FUNCTION_BLOCK FB_AxesEnable
VAR_INPUT
	bEnableAxes: 		BOOL := TRUE;
	bEnableXY:			BOOL;
	bEnableZp:			BOOL;
	bEnableZn:			BOOL;
	bReset:				BOOL;
	fOverride:			LREAL := 10;
END_VAR             	
VAR_OUTPUT          	
	bAllAxesReady:		BOOL := FALSE;
	fbError:			FB_Error;
END_VAR             	
VAR_IN_OUT          	
	stX:				AXIS_REF;
	stY:				AXIS_REF;
	stZ:				AXIS_REF;
END_VAR
VAR	
//Freigaben
	fbPowerX:			MC_Power;
	fbPowerY:			MC_Power;
	fbPowerZ:			MC_Power;
END_VAR


IF NOT (__ISVALIDREF(stX) AND __ISVALIDREF(stY) AND __ISVALIDREF(stZ)) THEN
	fbError.M_Set(1798, 'Üngültige Referenz der Achsen', 0, eID := E_ErrorIDs.eInvalidReference, eSrc := E_ErrorSrcs.ePlc);
	RETURN;
END_IF

IF bReset THEN
	fbError.M_Reset();
	bReset := FALSE;
END_IF

stX.ReadStatus();
stY.ReadStatus();
stZ.ReadStatus();

fbPowerX(
	Enable:=bEnableAxes AND bEnableXY, 
	Enable_Positive:=bEnableAxes AND bEnableXY, 
	Enable_Negative:=bEnableAxes AND bEnableXY, 
	Override:=fOverride, 
	BufferMode:= , 
	Axis:=stX, 
	Status=> , 
	Busy=> , 
	Active=> , 
	Error=> , 
	ErrorID=> );
	
fbPowerY(
	Enable:=bEnableAxes AND bEnableXY, 
	Enable_Positive:=bEnableAxes AND bEnableXY, 
	Enable_Negative:=bEnableAxes AND bEnableXY, 
	Override:=fOverride, 
	BufferMode:= , 
	Axis:=stY, 
	Status=> , 
	Busy=> , 
	Active=> , 
	Error=> , 
	ErrorID=> );	
	
fbPowerZ(
	Enable:=bEnableAxes, 
	Enable_Positive:=bEnableAxes AND bEnableZp, 
	Enable_Negative:=bEnableAxes AND bEnableZn, 
	Override:=fOverride, 
	BufferMode:= , 
	Axis:=stZ, 
	Status=> , 
	Busy=> , 
	Active=> , 
	Error=> , 
	ErrorID=> );		
	
bAllAxesReady := stX.Status.Operational AND stY.Status.Operational AND stZ.Status.Operational;
IF fbPowerX.Error THEN
	fbError.M_Set(fbPowerX.ErrorID, 'Achse X Error', 0, eID := E_ErrorIDs.eAxisRelease, eSrc := E_ErrorSrcs.eAxisX);
ELSIF fbPowerY.Error THEN
	fbError.M_Set(fbPowerY.ErrorID, 'Achse Y Error', 0, eID := E_ErrorIDs.eAxisRelease, eSrc := E_ErrorSrcs.eAxisY);
ELSIF fbPowerZ.Error THEN
	fbError.M_Set(fbPowerZ.ErrorID, 'Achse Z Error', 0, eID := E_ErrorIDs.eAxisRelease, eSrc := E_ErrorSrcs.eAxisZ);
END_IF

METHOD M_DisableAxes
VAR_INPUT
END_VAR
bEnableAxes:= FALSE;
bEnableXY:= FALSE;
bEnableZp:= FALSE; 
bEnableZn:= FALSE;
END_METHOD

METHOD M_EnableAxes
VAR_INPUT
END_VAR
bEnableAxes:= TRUE;
bEnableXY:= TRUE;
bEnableZp:= TRUE; 
bEnableZn:= TRUE;
END_METHOD

END_FUNCTION_BLOCK

(* stored: Version 1.1.0.1, ProductVersion 3.1.4024.12
   POU FB_AxesEnable: Id {99414854-69cd-49ca-984e-d64791bedf4d}, SpecialFunc None
   Method M_DisableAxes: Id {48de92bb-1aa1-4a25-8e68-a47f73eac763}
   Method M_EnableAxes: Id {14e6e14f-2c7a-408f-8812-95d47b4eda5b} *)
